SUBAPPLICATION Uebung_231 (* FIFO: Tastendruecke puffern, Q1 blinkt je Wert einmal (PROCESSED-Handshake) *)
  (* Standard: 61499-2; Description: Copyright (c) 2026 Meisterschulen am Ostbahnhof This program and the accompanying materials are made available under the terms of the Eclipse Public License 2.0 which is available at https://www.eclipse.org/legal/epl-2.0/ SPDX-License-Identifier: EPL-2.0 *)
  (* Version 1.0, 2026-11-08, Franz Höpfinger, Meisterschulen am Ostbahnhof, initial API and implementation and/or initial documentation *)
  PACKAGE Uebungen;
  IMPORT logiBUS::io::DI::logiBUS_DI::Input_I1;
  IMPORT logiBUS::io::DI::logiBUS_DI::Input_I4;
  IMPORT logiBUS::io::DI::logiBUS_DI_Events::BUTTON_SINGLE_CLICK;
  IMPORT logiBUS::io::DQ::logiBUS_DO::Output_Q1;
  IMPORT logiBUS::io::DQ::logiBUS_DO::Output_Q2;
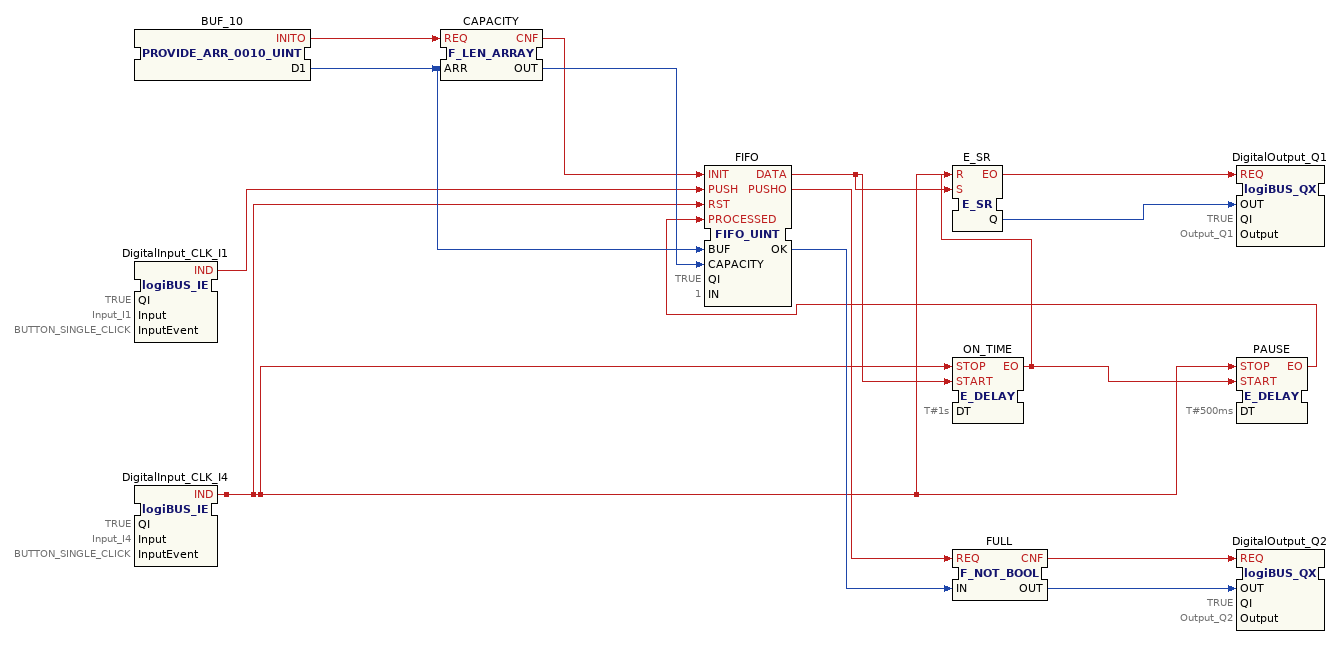
  FBS
    BUF_10 : eclipse4diac::convert::providers::PROVIDE_ARR_0010_UINT;
    CAPACITY : eclipse4diac::utils::arrays::F_LEN_ARRAY;
    FIFO : FIFO::FIFO_UINT(QI := TRUE, IN := 1);
    DigitalInput_CLK_I1 : logiBUS::io::DI::logiBUS_IE(QI := TRUE, Input := Input_I1, InputEvent := BUTTON_SINGLE_CLICK);
    DigitalInput_CLK_I4 : logiBUS::io::DI::logiBUS_IE(QI := TRUE, Input := Input_I4, InputEvent := BUTTON_SINGLE_CLICK);
    E_SR : iec61499::events::E_SR;
    ON_TIME : iec61499::events::E_DELAY(DT := T#1s);
    PAUSE : iec61499::events::E_DELAY(DT := T#500ms);
    DigitalOutput_Q1 : logiBUS::io::DQ::logiBUS_QX(QI := TRUE, Output := Output_Q1);
    FULL : iec61131::booleanOperators::F_NOT_BOOL;
    DigitalOutput_Q2 : logiBUS::io::DQ::logiBUS_QX(QI := TRUE, Output := Output_Q2);
  END_FBS
  EVENT_CONNECTIONS
    BUF_10.INITO TO CAPACITY.REQ;
    CAPACITY.CNF TO FIFO.INIT;
    DigitalInput_CLK_I1.IND TO FIFO.PUSH;
    DigitalInput_CLK_I4.IND TO FIFO.RST;
    DigitalInput_CLK_I4.IND TO ON_TIME.STOP;
    DigitalInput_CLK_I4.IND TO PAUSE.STOP;
    DigitalInput_CLK_I4.IND TO E_SR.R;
    FIFO.DATA TO E_SR.S;
    FIFO.DATA TO ON_TIME.START;
    ON_TIME.EO TO E_SR.R;
    ON_TIME.EO TO PAUSE.START;
    PAUSE.EO TO FIFO.PROCESSED;
    E_SR.EO TO DigitalOutput_Q1.REQ;
    FIFO.PUSHO TO FULL.REQ;
    FULL.CNF TO DigitalOutput_Q2.REQ;
  END_CONNECTIONS
  DATA_CONNECTIONS
    BUF_10.D1 TO CAPACITY.ARR;
    BUF_10.D1 TO FIFO.BUF;
    CAPACITY.OUT TO FIFO.CAPACITY;
    E_SR.Q TO DigitalOutput_Q1.OUT;
    FIFO.OK TO FULL.IN;
    FULL.OUT TO DigitalOutput_Q2.OUT;
  END_CONNECTIONS
END_SUBAPPLICATION
